# EPICS substitutions: b-55B2VNC/src/main/c++/nds3-6683h/src/main/epics/ndsNisyncApp/Db/nisyncDevice6683H-basic.substitutions
#State Machine for the device
file "nisync_Device.template" {
pattern
{
	BOARDTYPE,
	BOARDTYPEIDX,
	CBS1,
	CBS2
}

{
	"B",
	"0",
	"TEST",
	"FCT0"
}

}
# Firmware node
file "nisync_Firmware.template" {
pattern
{
	BOARDTYPE,
	BOARDTYPEIDX,
	CBS1,
	CBS2,
	FIRMWARE_NAME,
}

{
	"B",
	"0",
	"TEST",
	"FCT0",
	"Firm",
}

}

file "nisync_Routing.template" {
pattern
{
	BOARDTYPE,
	BOARDTYPEIDX,
	CBS1,
	CBS2,
	ROUTING_NAME
}

{
	"B",
	"0",
	"TEST",
	"FCT0",
	"Routing"
}

}
file "nisync_Timing.template" {
pattern
{
	BOARDTYPE,
	BOARDTYPEIDX,
	CBS1,
	CBS2,
	TIMING_NAME,
}

{
	"B",
	"0",
	"TEST",
	"FCT0",
	"Timing",
}

}
